Fanuc KAREL source: kt00508.KL

PROGRAM KT00508
%STACKSIZE=65535
%PRIORITY=65535
%NOLOCKGROUP
VAR
P1 : XYZWPR
P2 : JOINTPOS9
OUT : BOOLEAN
BEGIN
P1.X=1.0
-- UNRESOLVED_PC line 9 opcodes [49 7E 49 7E AC 23] marker_code=20
END KT00508
